(* IEC 61131-3 sources: Caravan/Archiv/12-04-19/Stations/MachineControl/MachineControl/Network/Power_Net, 1 file *)

(* ---- ONE_Power_Net_Table.st ---- *)
#define OBJECTS_CONFIG

FUNCTION GLOBAL TAB ONE_Power_Net
-1$UINT, 0$UINT,
0$UINT, 0$UINT,

2$UDINT,
TO_UDINT(357931502), "Battery_Class", 0$UINT, 0$UINT, 1$UINT,
TO_UDINT(1681589219), "Grid_Class", 0$UINT, 0$UINT, 1$UINT,

_NO_ATTR, TO_UDINT(3296425297), "BATTERY_CLASS1",

_NO_ATTR, TO_UDINT(3132843894), "GRID_CLASS1",

//Internal connections
0$UDINT,
0$UDINT,
0$UDINT,
0$UDINT,

//Initialization values
0$UDINT,
0$UDINT,

//Symbolic initialization values
0$UDINT,
0$UDINT,

//Initialization of string values
0$UDINT,
0$UDINT,

//Configuration of tasks (RealTime, Cyclic, Background)
0$UDINT,
0$UDINT,

0$UDINT,
2$UDINT,
TO_UDINT(0), (100)$UDINT, 4194303$DINT, 	//BATTERY_CLASS1
TO_UDINT(1), (50)$UDINT, 4194303$DINT, 	//GRID_CLASS1

0$UDINT,
0$UDINT,

//External connections
0$UDINT,
5$UDINT,
TO_UDINT(0), "ActualAmps1_C", C_DIR, TO_UDINT(3157766682), "AI0881","TMP_1",
TO_UDINT(0), "ActualAmps2_C", C_DIR, TO_UDINT(3157766682), "AI0881","TMP_2",
TO_UDINT(0), "ActualVoltage_C", C_DIR, TO_UDINT(46500714), "AI0751","AI4",
TO_UDINT(0), "ActualTowCarVoltage_C", C_DIR, TO_UDINT(46500714), "AI0751","AI6",
TO_UDINT(1), "ActualAmps_C", C_DIR, TO_UDINT(46500714), "AI0751","AI5",

//Magic internal connections
0$UDINT,
0$UDINT,

//Configuration of timeslots of tasks (RealTime, Cyclic)
#ifdef __LSLLDR_TIMESLOTS__
0$UDINT,
0$UDINT,

0$UDINT,
0$UDINT,

#endif //__LSLLDR_TIMESLOTS__

//MultiMaster connections
#ifdef __LSLLDR_MULTIMASTER__
0$UDINT,
0$UDINT,
#endif //__LSLLDR_MULTIMASTER__

//Configuration for task ID (RealTime, CyclicTime)
#ifdef __LSLLDR_TASKID__
"\\\\TASKS2  "
0$UDINT,
0$UDINT,

0$UDINT,
2$UDINT,
(0)$UDINT, 	//BATTERY_CLASS1
(0)$UDINT, 	//GRID_CLASS1

0$UDINT,
0$UDINT,

#endif //__LSLLDR_TASKID__

END_FUNCTION
